(* IEC 61131-3 sources: plc-patterns-examples/listings/BottleFiller, 39 files *)

(* ---- E_ActuatorTarget.st ---- *)
{attribute 'qualified_only'}
{attribute 'strict'}
{attribute 'to_string'}
TYPE E_ActuatorTarget :
(
    None      := 0,     // no move commanded yet; what the outputs do is up to the actuator
    Extended  := 10,
    Retracted := 20
);
END_TYPE

(* ---- E_DeviceSource.st ---- *)
{attribute 'qualified_only'}
{attribute 'strict'}
{attribute 'to_string'}
TYPE E_DeviceSource :
(
    Undefined       := 0,
    FinalHardware   := 1,
    SimilarHardware := 2,
    Simulation      := 3,
    Test            := 4
);
END_TYPE

(* ---- E_FillStep.st ---- *)
{attribute 'qualified_only'}
{attribute 'strict'}
{attribute 'to_string'}
TYPE E_FillStep :
(
    Undefined := 0,
    Idle      := 10,
    Opening   := 20,
    Filling   := 30,
    Closing   := 40,
    Done      := 50,
    Error     := 900
);
END_TYPE

(* ---- E_LineState.st ---- *)
{attribute 'qualified_only'}
{attribute 'strict'}
{attribute 'to_string'}
TYPE E_LineState :
(
    Stopped      := 0,
    Filling      := 10,
    Transferring := 20,
    Faulted      := 900
);
END_TYPE

(* ---- E_OperationState.st ---- *)
{attribute 'qualified_only'}
{attribute 'strict'}
{attribute 'to_string'}
TYPE E_OperationState :
(
    Idle  := 0,     // never started
    Busy  := 1,
    Done  := 2,
    Error := 3
);
END_TYPE

(* ---- E_PickStep.st ---- *)
{attribute 'qualified_only'}
{attribute 'strict'}
{attribute 'to_string'}
TYPE E_PickStep :
(
    Undefined      := 0,
    Idle           := 10,
    LowerToPick    := 20,
    Grip           := 30,
    RaiseWithPart  := 40,
    SlideOut       := 50,
    LowerToPlace   := 60,
    ClampPart      := 65,
    OpenGripper    := 70,
    RaiseEmpty     := 80,
    ReleaseFixture := 85,
    SlideIn        := 90,
    Done           := 100,
    Error          := 900
);
END_TYPE

(* ---- GVL_Hmi.st ---- *)
{attribute 'qualified_only'}
VAR_GLOBAL
    // From the HMI
    StartButton      : BOOL;
    StopButton       : BOOL;
    ResetButton      : BOOL;

    // To the HMI
    LineState        : E_LineState;
    IsStopping       : BOOL;
    FaultText        : STRING;
    NotFinalDevices  : STRING(255);         // every device that isn't the machine's own; empty on the machine
END_VAR

(* ---- GVL_Io.st ---- *)
{attribute 'qualified_only'}
VAR_GLOBAL
    // Filling station
    TankValveCoil  AT %Q* : BOOL;
    TankValveOpen  AT %I* : BOOL;
    DrainValveCoil AT %Q* : BOOL;
    DrainValveOpen AT %I* : BOOL;
    TankLevel      AT %I* : DINT;           // level sensor process data, 0.1 mm
    TankSensorOk   AT %I* : BOOL;           // the sensor's valid bit; see the project document

    // Pick-and-place station
    LiftValve      AT %Q* : BOOL;
    LiftDown       AT %I* : BOOL;
    LiftUp         AT %I* : BOOL;
    SlideOutCoil   AT %Q* : BOOL;
    SlideInCoil    AT %Q* : BOOL;
    SlideOut       AT %I* : BOOL;
    SlideIn        AT %I* : BOOL;
    GripperValve   AT %Q* : BOOL;
    GripperClosed  AT %I* : BOOL;
    GripperOpen    AT %I* : BOOL;
END_VAR

(* ---- GVL_Sim.st ---- *)
{attribute 'qualified_only'}
VAR_GLOBAL
    // Failure hooks for the simulated devices, set from the HMI or a watch
    // window. Each one acts only while its device is simulated.
    TankValveStuck  : BOOL;
    DrainValveStuck : BOOL;
    LiftStuck       : BOOL;
    SlideStuck      : BOOL;
    GripperStuck    : BOOL;
END_VAR

(* ---- GVL_Site.st ---- *)
{attribute 'qualified_only'}
VAR_GLOBAL CONSTANT
    // Edited for each controller; a release never overwrites this list.
    // FinalHardware on the machine. As delivered, everything is simulated.
    TankValveSource  : E_DeviceSource := E_DeviceSource.Simulation;
    DrainValveSource : E_DeviceSource := E_DeviceSource.Simulation;
    TankLevelSource  : E_DeviceSource := E_DeviceSource.Simulation;
    LiftSource       : E_DeviceSource := E_DeviceSource.Simulation;
    SlideSource      : E_DeviceSource := E_DeviceSource.Simulation;
    GripperSource    : E_DeviceSource := E_DeviceSource.Simulation;
    IsOnMachine      : BOOL := FALSE;   // TRUE on the real machine: anything not final is a fault
END_VAR

(* ---- ActuatorBase.st ---- *)
FUNCTION_BLOCK ABSTRACT ActuatorBase IMPLEMENTS I_Actuator, I_Cyclic
VAR
    _Name         : STRING(32);
    _MoveTimeout  : TIME := T#2S;
    _Target       : E_ActuatorTarget;
    _IsInPosition : BOOL;
    _HasFault     : BOOL;
    _FaultText    : STRING(80);
    _MoveTimer    : TON;
    _SettleTimer  : TON;
END_VAR
(*
    ActuatorBase

    The move-and-supervise skeleton shared by every actuator. CyclicLogic() is
    the template: it drives toward the target, checks arrival, supervises the
    move time, goes safe on a fault and lets the actuator settle.

    Derived blocks implement IsWired, DriveOutputs, IsAtPosition and DriveSafe,
    may override SettleTime, and call Configure() from their FB_init.
*)

METHOD PUBLIC FINAL CyclicLogic
// Not wired: report it, touch nothing
IF NOT IsWired() THEN
    _HasFault := TRUE;
    _FaultText := 'I/O not wired';
    RETURN;
END_IF

// Faulted: only the safe outputs, until Reset()
IF _HasFault THEN
    DriveSafe();
    RETURN;
END_IF

// Drive toward the target, and check whether it has arrived
DriveOutputs(Target := _Target);
_IsInPosition := IsAtPosition(Position := _Target);

// Supervise the move: the same rule for every actuator
_MoveTimer(IN := (_Target <> E_ActuatorTarget.None) AND NOT _IsInPosition, PT := _MoveTimeout);
IF _MoveTimer.Q THEN
    _HasFault := TRUE;
    _FaultText := 'Move did not finish in time';
    DriveSafe();
    RETURN;
END_IF

// Let it settle before reporting the position
_SettleTimer(IN := _IsInPosition, PT := SettleTime);

METHOD PROTECTED ABSTRACT IsWired : BOOL

METHOD PROTECTED ABSTRACT DriveOutputs
VAR_INPUT
    Target : E_ActuatorTarget;
END_VAR

METHOD PROTECTED ABSTRACT IsAtPosition : BOOL
VAR_INPUT
    Position : E_ActuatorTarget;
END_VAR

METHOD PROTECTED ABSTRACT DriveSafe

PROPERTY PROTECTED SettleTime : TIME
GET: SettleTime := T#0S;           // most actuators report as soon as the sensor confirms

METHOD PROTECTED Configure
VAR_INPUT
    Name        : STRING(32);
    MoveTimeout : TIME;
END_VAR
_Name := Name;
_MoveTimeout := MoveTimeout;

METHOD PUBLIC Extend
MoveTo(Target := E_ActuatorTarget.Extended);

METHOD PUBLIC Retract
MoveTo(Target := E_ActuatorTarget.Retracted);

METHOD PRIVATE MoveTo
VAR_INPUT
    Target : E_ActuatorTarget;
END_VAR
IF _HasFault OR Target = _Target THEN
    RETURN;                        // faulted: Reset() first. Same target: keep the move running.
END_IF
_Target := Target;
_MoveTimer(IN := FALSE);           // every new move gets the full timeout
_SettleTimer(IN := FALSE);

METHOD PUBLIC Reset
_HasFault := FALSE;
_FaultText := '';
_Target := E_ActuatorTarget.None;
_MoveTimer(IN := FALSE);
_SettleTimer(IN := FALSE);

PROPERTY PUBLIC IsExtended : BOOL
GET: IsExtended := NOT _HasFault AND _Target = E_ActuatorTarget.Extended AND _SettleTimer.Q;

PROPERTY PUBLIC IsRetracted : BOOL
GET: IsRetracted := NOT _HasFault AND _Target = E_ActuatorTarget.Retracted AND _SettleTimer.Q;

PROPERTY PUBLIC HasFault : BOOL
GET: HasFault := _HasFault;

PROPERTY PUBLIC FaultText : STRING
GET: FaultText := _FaultText;

PROPERTY PUBLIC Name : STRING
GET: Name := _Name;

(* ---- ActuatorRouter.st ---- *)
FUNCTION_BLOCK ActuatorRouter IMPLEMENTS I_Actuator, I_Cyclic
VAR
    _Name   : STRING(32);
    _Source : E_DeviceSource;
    _Chosen : I_Actuator;
END_VAR
(*
    ActuatorRouter

    One I_Actuator in front of up to four candidates, chosen once by the
    site setting. Only the chosen candidate is run. A source with no
    candidate (0) is never at either end, and reports a fault.
*)

METHOD FB_init : BOOL
VAR_INPUT
    bInitRetains    : BOOL;
    bInCopyCode     : BOOL;
    Name            : STRING(32);
    Source          : E_DeviceSource;
    FinalHardware   : I_Actuator;
    SimilarHardware : I_Actuator;
    Simulation      : I_Actuator;
    Test            : I_Actuator;
END_VAR
_Name := Name;
_Source := Source;
CASE Source OF
    E_DeviceSource.FinalHardware:   _Chosen := FinalHardware;
    E_DeviceSource.SimilarHardware: _Chosen := SimilarHardware;
    E_DeviceSource.Simulation:      _Chosen := Simulation;
    E_DeviceSource.Test:            _Chosen := Test;
END_CASE

METHOD PUBLIC CyclicLogic
VAR
    Cyclic : I_Cyclic;
END_VAR
IF _Chosen <> 0 AND_THEN __QUERYINTERFACE(_Chosen, Cyclic) THEN
    Cyclic.CyclicLogic();              // only the chosen candidate runs
END_IF

METHOD PUBLIC Extend
IF _Chosen <> 0 THEN
    _Chosen.Extend();
END_IF

METHOD PUBLIC Retract
IF _Chosen <> 0 THEN
    _Chosen.Retract();
END_IF

METHOD PUBLIC Reset
IF _Chosen <> 0 THEN
    _Chosen.Reset();
END_IF

PROPERTY PUBLIC IsExtended : BOOL
GET: IsExtended := _Chosen <> 0 AND_THEN _Chosen.IsExtended;

PROPERTY PUBLIC IsRetracted : BOOL
GET: IsRetracted := _Chosen <> 0 AND_THEN _Chosen.IsRetracted;

PROPERTY PUBLIC Name : STRING
GET: Name := _Name;

PROPERTY PUBLIC HasFault : BOOL
GET: HasFault := _Chosen = 0 OR_ELSE _Chosen.HasFault;

PROPERTY PUBLIC FaultText : STRING
GET:
IF _Chosen = 0 THEN
    FaultText := 'No device for this source';
ELSE
    FaultText := _Chosen.FaultText;
END_IF

PROPERTY PUBLIC Source : E_DeviceSource
GET: Source := _Source;

(* ---- DoubleSolenoidCylinder.st ---- *)
FUNCTION_BLOCK DoubleSolenoidCylinder EXTENDS ActuatorBase
VAR
    _ExtendCoil      : REFERENCE TO BOOL;
    _RetractCoil     : REFERENCE TO BOOL;
    _ExtendedSensor  : REFERENCE TO BOOL;
    _RetractedSensor : REFERENCE TO BOOL;
END_VAR
(*
    DoubleSolenoidCylinder

    One coil per direction. With both coils off, the valve holds the cylinder
    where it is. An end sensor at each end.
*)

METHOD FB_init : BOOL
VAR_INPUT
    bInitRetains    : BOOL;
    bInCopyCode     : BOOL;
    Name            : STRING(32);
    MoveTimeout     : TIME;
    ExtendCoil      : REFERENCE TO BOOL;
    RetractCoil     : REFERENCE TO BOOL;
    ExtendedSensor  : REFERENCE TO BOOL;
    RetractedSensor : REFERENCE TO BOOL;
END_VAR
_ExtendCoil REF= ExtendCoil;
_RetractCoil REF= RetractCoil;
_ExtendedSensor REF= ExtendedSensor;
_RetractedSensor REF= RetractedSensor;
Configure(Name := Name, MoveTimeout := MoveTimeout);

METHOD PROTECTED IsWired : BOOL
IsWired := __ISVALIDREF(_ExtendCoil) AND __ISVALIDREF(_RetractCoil)
       AND __ISVALIDREF(_ExtendedSensor) AND __ISVALIDREF(_RetractedSensor);

METHOD PROTECTED DriveOutputs
VAR_INPUT
    Target : E_ActuatorTarget;
END_VAR
_ExtendCoil := Target = E_ActuatorTarget.Extended;
_RetractCoil := Target = E_ActuatorTarget.Retracted;  // None: both off, so it holds

METHOD PROTECTED IsAtPosition : BOOL
VAR_INPUT
    Position : E_ActuatorTarget;
END_VAR
CASE Position OF
    E_ActuatorTarget.Extended:
        IsAtPosition := _ExtendedSensor AND NOT _RetractedSensor;
    E_ActuatorTarget.Retracted:
        IsAtPosition := _RetractedSensor AND NOT _ExtendedSensor;
ELSE
    IsAtPosition := FALSE;
END_CASE

METHOD PROTECTED DriveSafe
_ExtendCoil := FALSE;                               // both off: the cylinder stays where it is
_RetractCoil := FALSE;

(* ---- DrainTankCommand.st ---- *)
FUNCTION_BLOCK DrainTankCommand IMPLEMENTS I_Command
VAR CONSTANT
    EmptyLevel : REAL := 2.0;          // percent
END_VAR
VAR
    _DrainValve   : I_FillValve;
    _Level        : I_LevelSensor;
    _Clock        : I_Clock;
    _Timeout      : LTIME;
    _StartedAt    : LTIME;
    _State        : E_OperationState;
    _FaultText    : STRING;
    _IsConfigured : BOOL;
END_VAR
(*
    DrainTankCommand

    Opens the drain valve until the tank reads empty. Ends in Error if the
    level sensor is invalid, the valve faults, or the tank isn't empty
    within the timeout. Every ending closes the drain valve.
*)

METHOD FB_init : BOOL
VAR_INPUT
    bInitRetains : BOOL;
    bInCopyCode  : BOOL;
    DrainValve   : I_FillValve;     // any on/off valve with feedback fits this contract
    Level        : I_LevelSensor;
    Clock        : I_Clock;
    Timeout      : LTIME;
END_VAR
_DrainValve := DrainValve;
_Level := Level;
_Clock := Clock;
_Timeout := Timeout;
_IsConfigured := DrainValve <> 0 AND Level <> 0 AND Clock <> 0;

METHOD PUBLIC Start
IF _State = E_OperationState.Busy THEN
    RETURN;
END_IF
IF NOT _IsConfigured THEN
    _State := E_OperationState.Error;
    _FaultText := 'Drain command not wired';
    RETURN;
END_IF
_StartedAt := _Clock.Now;
_FaultText := '';
_State := E_OperationState.Busy;
_DrainValve.Open();

METHOD PUBLIC CyclicLogic
IF _State <> E_OperationState.Busy THEN
    RETURN;
END_IF

IF NOT _Level.IsValid THEN
    Finish(Outcome := E_OperationState.Error, Text := 'Level sensor invalid');
ELSIF _DrainValve.HasFault THEN
    Finish(Outcome := E_OperationState.Error, Text := _DrainValve.FaultText);
ELSIF _Level.Level <= EmptyLevel THEN
    Finish(Outcome := E_OperationState.Done, Text := '');
ELSIF _Clock.Now - _StartedAt >= _Timeout THEN
    Finish(Outcome := E_OperationState.Error, Text := 'Tank did not empty in time');
END_IF

METHOD PUBLIC Abort
IF _State = E_OperationState.Busy THEN
    Finish(Outcome := E_OperationState.Error, Text := 'Aborted');
END_IF

METHOD PRIVATE Finish
VAR_INPUT
    Outcome : E_OperationState;
    Text    : STRING;
END_VAR
_DrainValve.Close();                 // every ending, good or bad, leaves the drain closed
_State := Outcome;
_FaultText := Text;

PROPERTY PUBLIC Name : STRING
GET: Name := 'Drain tank';

PROPERTY PUBLIC State : E_OperationState
GET: State := _State;

PROPERTY PUBLIC FaultText : STRING
GET: FaultText := _FaultText;

(* ---- EquipmentGroup.st ---- *)
FUNCTION_BLOCK EquipmentGroup IMPLEMENTS I_Diagnosable, I_Resettable
VAR CONSTANT
    MaxChildren : DINT := 16;
END_VAR
VAR
    _Name        : STRING(32);
    _Children    : ARRAY[0..MaxChildren - 1] OF I_Diagnosable;
    _Resettables : ARRAY[0..MaxChildren - 1] OF I_Resettable;
    _Count       : DINT;
END_VAR
(*
    EquipmentGroup

    A named group of devices or other groups, behind the same interfaces
    as one device. It has a fault while any child has one, and reports
    the first faulted child's text, prefixed with that child's name.
    Reset() resets every child that implements I_Resettable.
    AddChild() is called while wiring, before the group is first asked.
*)

METHOD FB_init : BOOL
VAR_INPUT
    bInitRetains : BOOL;
    bInCopyCode  : BOOL;
    Name         : STRING(32);
END_VAR
_Name := Name;

METHOD PUBLIC AddChild : BOOL
VAR_INPUT
    Child : I_Diagnosable;
END_VAR
VAR
    Me         : I_Diagnosable;
    Resettable : I_Resettable;
    i          : DINT;
END_VAR
Me := THIS^;
IF Child = 0 OR Child = Me OR _Count >= MaxChildren THEN
    AddChild := FALSE;
    RETURN;
END_IF
FOR i := 0 TO _Count - 1 DO           // the same child only once
    IF _Children[i] = Child THEN
        AddChild := FALSE;
        RETURN;
    END_IF
END_FOR
_Children[_Count] := Child;
IF __QUERYINTERFACE(Child, Resettable) THEN
    _Resettables[_Count] := Resettable;
END_IF
_Count := _Count + 1;
AddChild := TRUE;

METHOD PUBLIC Reset
VAR
    i : DINT;
END_VAR
FOR i := 0 TO _Count - 1 DO
    IF _Resettables[i] <> 0 THEN
        _Resettables[i].Reset();
    END_IF
END_FOR

METHOD PRIVATE FirstFaultIndex : DINT
VAR
    i : DINT;
END_VAR
FOR i := 0 TO _Count - 1 DO
    IF _Children[i].HasFault THEN
        FirstFaultIndex := i;
        RETURN;
    END_IF
END_FOR
FirstFaultIndex := _Count;            // no child has a fault

METHOD PRIVATE DescribeFault : STRING
VAR_INPUT
    Index : DINT;
END_VAR
IF Index < _Count THEN
    DescribeFault := CONCAT(CONCAT(_Children[Index].Name, ': '), _Children[Index].FaultText);
END_IF

PROPERTY PUBLIC Name : STRING
GET: Name := _Name;

PROPERTY PUBLIC HasFault : BOOL
GET: HasFault := FirstFaultIndex() < _Count;

PROPERTY PUBLIC FaultText : STRING
GET: FaultText := DescribeFault(Index := FirstFaultIndex());

PROPERTY PUBLIC ChildCount : DINT
GET: ChildCount := _Count;

(* ---- FakeClock.st ---- *)
FUNCTION_BLOCK FakeClock IMPLEMENTS I_Clock
VAR
    _Now : LTIME;
END_VAR
(*
    FakeClock

    Stands still until the test moves it.
*)

METHOD PUBLIC Advance
VAR_INPUT
    Duration : LTIME;
END_VAR
_Now := _Now + Duration;

PROPERTY PUBLIC Now : LTIME
GET: Now := _Now;

(* ---- FakeEquipmentModule.st ---- *)
FUNCTION_BLOCK FakeEquipmentModule IMPLEMENTS I_EquipmentModule, I_Resettable
VAR
    _Name        : STRING(32);
    _IsCycleDone : BOOL;
    _HasFault    : BOOL;
    _StartCount  : DINT;
    _ResetCount  : DINT;
END_VAR
(*
    FakeEquipmentModule

    Test double for I_EquipmentModule. Counts the cycles it was asked for
    and the resets it received. A requested cycle finishes when the test
    calls FinishCycle(); a fault is reported while the test sets one.
*)

METHOD FB_init : BOOL
VAR_INPUT
    bInitRetains : BOOL;
    bInCopyCode  : BOOL;
    Name         : STRING(32);
END_VAR
_Name := Name;

METHOD PUBLIC StartCycle
_StartCount := _StartCount + 1;
_IsCycleDone := FALSE;

METHOD PUBLIC Reset
_ResetCount := _ResetCount + 1;

METHOD PUBLIC FinishCycle
_IsCycleDone := TRUE;

METHOD PUBLIC SetFault
VAR_INPUT
    IsActive : BOOL;
END_VAR
_HasFault := IsActive;

PROPERTY PUBLIC Name : STRING
GET: Name := _Name;

PROPERTY PUBLIC HasFault : BOOL
GET: HasFault := _HasFault;

PROPERTY PUBLIC FaultText : STRING
GET:
IF _HasFault THEN
    FaultText := 'Simulated fault';
ELSE
    FaultText := '';
END_IF

PROPERTY PUBLIC IsCycleDone : BOOL
GET: IsCycleDone := _IsCycleDone;

PROPERTY PUBLIC StartCount : DINT
GET: StartCount := _StartCount;

PROPERTY PUBLIC ResetCount : DINT
GET: ResetCount := _ResetCount;

(* ---- FieldbusLevelSensor.st ---- *)
FUNCTION_BLOCK FieldbusLevelSensor IMPLEMENTS I_LevelSensor
VAR
    _FieldbusLevel     : REFERENCE TO DINT;
    _IsCommunicationOk : REFERENCE TO BOOL;
    _TankHeight        : REAL;
    _IsConfigured      : BOOL;
END_VAR
(* FieldbusLevelSensor: a level sensor that reports its reading over a fieldbus, in 0.1 mm. *)

METHOD FB_init : BOOL
VAR_INPUT
    bInitRetains      : BOOL;
    bInCopyCode       : BOOL;
    FieldbusLevel     : REFERENCE TO DINT;   // process data from the sensor, 0.1 mm
    IsCommunicationOk : REFERENCE TO BOOL;
    TankHeight        : REAL;                // mm
END_VAR
_FieldbusLevel REF= FieldbusLevel;
_IsCommunicationOk REF= IsCommunicationOk;
_TankHeight := TankHeight;
_IsConfigured := __ISVALIDREF(FieldbusLevel) AND __ISVALIDREF(IsCommunicationOk) AND TankHeight > 0.0;

PROPERTY PUBLIC IsValid : BOOL
GET: IsValid := _IsConfigured AND_THEN _IsCommunicationOk;

PROPERTY PUBLIC Level : REAL
GET:
IF IsValid THEN
    Level := LIMIT(0.0, DINT_TO_REAL(_FieldbusLevel) / 10.0 / _TankHeight * 100.0, 100.0);
ELSE
    Level := 0.0;
END_IF

(* ---- FillingModule.st ---- *)
FUNCTION_BLOCK FillingModule EXTENDS ModuleGroup IMPLEMENTS I_EquipmentModule
VAR
    _Fill             : REFERENCE TO FillSequence;
    _Dose             : I_Command;
    _IsCycleRequested : BOOL;
    _IsFilling        : BOOL;
    _IsDosing         : BOOL;
    _HasDoseFault     : BOOL;
    _DoseFault        : STRING;
    _IsConfigured     : BOOL;
END_VAR
(*
    FillingModule

    The filling station. One cycle measures one dose: the fill sequence
    fills the dosing tank to its target level, then the dose command
    drains it into the bottle below. Runs both before its valves. It has
    a fault while a valve has one, the fill sequence has stopped with an
    error, or the last dose ended in Error; Reset() clears all three.
*)

METHOD FB_init : BOOL
VAR_INPUT
    bInitRetains : BOOL;
    bInCopyCode  : BOOL;
    Name         : STRING(32);                  // for EquipmentGroup
    Fill         : REFERENCE TO FillSequence;
    Dose         : I_Command;
END_VAR
_Fill REF= Fill;
_Dose := Dose;
_IsConfigured := __ISVALIDREF(Fill) AND Dose <> 0;

METHOD PUBLIC StartCycle
_IsCycleRequested := TRUE;

METHOD PROTECTED BeforeChildren
IF NOT _IsConfigured THEN
    RETURN;
END_IF

// A new cycle starts with the fill, once the station is free
IF _IsCycleRequested AND NOT _IsFilling AND NOT _IsDosing
   AND (_Fill.CurrentStep = E_FillStep.Idle OR _Fill.CurrentStep = E_FillStep.Done) THEN
    _Fill.Start();
    _IsFilling := TRUE;
    _IsCycleRequested := FALSE;
END_IF
_Fill.CyclicLogic();

// The tank is at its level: dose it into the bottle
IF _IsFilling AND _Fill.IsDone THEN
    _IsFilling := FALSE;
    _Dose.Start();
    _IsDosing := TRUE;
END_IF
IF _IsDosing THEN
    _Dose.CyclicLogic();
    IF _Dose.State = E_OperationState.Error THEN
        _HasDoseFault := TRUE;
        _DoseFault := _Dose.FaultText;
        _IsDosing := FALSE;
    ELSIF _Dose.State = E_OperationState.Done THEN
        _IsDosing := FALSE;
    END_IF
END_IF

METHOD PUBLIC Reset
SUPER^.Reset();                                 // the valves
IF NOT _IsConfigured THEN
    RETURN;
END_IF
_Fill.Reset();
IF _IsDosing THEN
    _Dose.Abort();                              // closes the drain valve
END_IF
_IsCycleRequested := FALSE;
_IsFilling := FALSE;
_IsDosing := FALSE;
_HasDoseFault := FALSE;
_DoseFault := '';

PROPERTY PUBLIC IsCycleDone : BOOL
GET:
IsCycleDone := _IsConfigured AND_THEN (NOT _IsCycleRequested AND NOT _IsFilling AND NOT _IsDosing
                                             AND _Dose.State = E_OperationState.Done);

PROPERTY PUBLIC HasFault : BOOL
GET:
IF NOT _IsConfigured THEN
    HasFault := TRUE;
ELSE
    HasFault := SUPER^.HasFault OR _Fill.HasError OR _HasDoseFault;
END_IF

PROPERTY PUBLIC FaultText : STRING
GET:
IF NOT _IsConfigured THEN
    FaultText := 'Filling station not wired';
ELSIF SUPER^.HasFault THEN
    FaultText := SUPER^.FaultText;              // the valve, by name
ELSIF _Fill.HasError THEN
    FaultText := 'Fill stopped; reset to continue';
ELSIF _HasDoseFault THEN
    FaultText := CONCAT('Dose: ', _DoseFault);
ELSE
    FaultText := '';
END_IF

(* ---- FillSequence.st ---- *)
FUNCTION_BLOCK FillSequence
VAR
    _LevelSensor      : I_LevelSensor;
    _FillValve        : I_FillValve;
    _TargetLevel      : REAL := 80.0;
    _CurrentStep      : E_FillStep := E_FillStep.Idle;
    _IsStartRequested : BOOL;
    _IsResetRequested : BOOL;
    _IsConfigured     : BOOL;
END_VAR
(*
    FillSequence

    Opens the fill valve, waits for the target level, closes the valve.
    Talks only to I_LevelSensor and I_FillValve, injected through FB_init.

    Call CyclicLogic() once per cycle. Start() and Reset() are requests,
    seen during the next CyclicLogic() call.
*)

METHOD PUBLIC Start
_IsStartRequested := TRUE;

METHOD PUBLIC Reset
_IsResetRequested := TRUE;

METHOD PUBLIC CyclicLogic
IF NOT _IsConfigured THEN
    _CurrentStep := E_FillStep.Error;   // not wired: fail safe, never call through 0
    RETURN;
END_IF

CASE _CurrentStep OF
    E_FillStep.Idle, E_FillStep.Done:
        IF _IsStartRequested THEN
            _CurrentStep := E_FillStep.Opening;
        END_IF

    E_FillStep.Opening:
        _FillValve.Open();
        IF _FillValve.IsOpen THEN
            _CurrentStep := E_FillStep.Filling;
        ELSIF _FillValve.HasFault THEN
            _CurrentStep := E_FillStep.Error;
        END_IF

    E_FillStep.Filling:
        IF NOT _LevelSensor.IsValid OR _FillValve.HasFault THEN
            _CurrentStep := E_FillStep.Error;
        ELSIF _LevelSensor.Level >= _TargetLevel THEN
            _CurrentStep := E_FillStep.Closing;
        END_IF

    E_FillStep.Closing:
        _FillValve.Close();
        IF _FillValve.IsClosed THEN
            _CurrentStep := E_FillStep.Done;
        ELSIF _FillValve.HasFault THEN
            _CurrentStep := E_FillStep.Error;
        END_IF

    E_FillStep.Error:
        _FillValve.Close();             // the one promise every valve keeps
        IF _IsResetRequested AND _FillValve.IsClosed THEN
            _CurrentStep := E_FillStep.Idle;
        END_IF
END_CASE

_IsStartRequested := FALSE;
_IsResetRequested := FALSE;

PROPERTY PUBLIC TargetLevel : REAL
GET: TargetLevel := _TargetLevel;
SET: _TargetLevel := LIMIT(0.0, TargetLevel, 100.0);

PROPERTY PUBLIC CurrentStep : E_FillStep
GET: CurrentStep := _CurrentStep;

PROPERTY PUBLIC IsBusy : BOOL
GET:
IsBusy := _CurrentStep = E_FillStep.Opening
            OR _CurrentStep = E_FillStep.Filling
            OR _CurrentStep = E_FillStep.Closing;

PROPERTY PUBLIC IsDone : BOOL
GET: IsDone := _CurrentStep = E_FillStep.Done;

PROPERTY PUBLIC HasError : BOOL
GET: HasError := _CurrentStep = E_FillStep.Error;

METHOD FB_init : BOOL
VAR_INPUT
    bInitRetains : BOOL;
    bInCopyCode  : BOOL;
    LevelSensor  : I_LevelSensor;
    FillValve    : I_FillValve;
END_VAR
_LevelSensor := LevelSensor;
_FillValve := FillValve;
_IsConfigured := LevelSensor <> 0 AND FillValve <> 0;   // stored: FB_init's return value is ignored

(* ---- FillValveRouter.st ---- *)
FUNCTION_BLOCK FillValveRouter IMPLEMENTS I_FillValve, I_Cyclic
VAR
    _Name   : STRING(32);
    _Source : E_DeviceSource;
    _Chosen : I_FillValve;
END_VAR
(*
    FillValveRouter

    One I_FillValve in front of up to four candidates. The site setting,
    given once in FB_init, chooses which candidate answers and which one
    is run. A source with no candidate (0) reports a fault and is never
    open.
*)

METHOD FB_init : BOOL
VAR_INPUT
    bInitRetains    : BOOL;
    bInCopyCode     : BOOL;
    Name            : STRING(32);
    Source          : E_DeviceSource;
    FinalHardware   : I_FillValve;
    SimilarHardware : I_FillValve;
    Simulation      : I_FillValve;
    Test            : I_FillValve;
END_VAR
_Name := Name;
_Source := Source;
CASE Source OF
    E_DeviceSource.FinalHardware:   _Chosen := FinalHardware;
    E_DeviceSource.SimilarHardware: _Chosen := SimilarHardware;
    E_DeviceSource.Simulation:      _Chosen := Simulation;
    E_DeviceSource.Test:            _Chosen := Test;
END_CASE

METHOD PUBLIC CyclicLogic
VAR
    Cyclic : I_Cyclic;
END_VAR
IF _Chosen <> 0 AND_THEN __QUERYINTERFACE(_Chosen, Cyclic) THEN
    Cyclic.CyclicLogic();              // only the chosen candidate runs
END_IF

METHOD PUBLIC Open
IF _Chosen <> 0 THEN
    _Chosen.Open();
END_IF

METHOD PUBLIC Close
IF _Chosen <> 0 THEN
    _Chosen.Close();
END_IF

PROPERTY PUBLIC IsOpen : BOOL
GET: IsOpen := _Chosen <> 0 AND_THEN _Chosen.IsOpen;

PROPERTY PUBLIC IsClosed : BOOL
GET: IsClosed := _Chosen <> 0 AND_THEN _Chosen.IsClosed;

PROPERTY PUBLIC Name : STRING
GET: Name := _Name;

PROPERTY PUBLIC HasFault : BOOL
GET: HasFault := _Chosen = 0 OR_ELSE _Chosen.HasFault;

PROPERTY PUBLIC FaultText : STRING
GET:
IF _Chosen = 0 THEN
    FaultText := 'No device for this source';
ELSE
    FaultText := _Chosen.FaultText;
END_IF

PROPERTY PUBLIC Source : E_DeviceSource
GET: Source := _Source;

(* ---- LevelSensorRouter.st ---- *)
FUNCTION_BLOCK LevelSensorRouter IMPLEMENTS I_LevelSensor, I_Cyclic
VAR
    _Name   : STRING(32);
    _Source : E_DeviceSource;
    _Chosen : I_LevelSensor;
END_VAR
(*
    LevelSensorRouter

    One I_LevelSensor in front of up to four candidates, chosen once by
    the site setting. A source with no candidate (0) is never valid.
*)

METHOD FB_init : BOOL
VAR_INPUT
    bInitRetains    : BOOL;
    bInCopyCode     : BOOL;
    Name            : STRING(32);
    Source          : E_DeviceSource;
    FinalHardware   : I_LevelSensor;
    SimilarHardware : I_LevelSensor;
    Simulation      : I_LevelSensor;
    Test            : I_LevelSensor;
END_VAR
_Name := Name;
_Source := Source;
CASE Source OF
    E_DeviceSource.FinalHardware:   _Chosen := FinalHardware;
    E_DeviceSource.SimilarHardware: _Chosen := SimilarHardware;
    E_DeviceSource.Simulation:      _Chosen := Simulation;
    E_DeviceSource.Test:            _Chosen := Test;
END_CASE

METHOD PUBLIC CyclicLogic
VAR
    Cyclic : I_Cyclic;
END_VAR
IF _Chosen <> 0 AND_THEN __QUERYINTERFACE(_Chosen, Cyclic) THEN
    Cyclic.CyclicLogic();              // only the chosen candidate runs
END_IF

PROPERTY PUBLIC Level : REAL
GET:
IF _Chosen <> 0 THEN
    Level := _Chosen.Level;
ELSE
    Level := 0.0;
END_IF

PROPERTY PUBLIC IsValid : BOOL
GET: IsValid := _Chosen <> 0 AND_THEN _Chosen.IsValid;

PROPERTY PUBLIC Name : STRING
GET: Name := _Name;

PROPERTY PUBLIC Source : E_DeviceSource
GET: Source := _Source;

(* ---- LineModule.st ---- *)
FUNCTION_BLOCK LineModule EXTENDS ModuleGroup
VAR
    _Filler           : I_EquipmentModule;
    _Transfer         : I_EquipmentModule;
    _State            : E_LineState;
    _IsStartRequested : BOOL;
    _IsStopping       : BOOL;
    _IsConfigured     : BOOL;
END_VAR
(*
    LineModule

    The machine module. Fills a bottle, moves it out, and repeats until
    stopped. Commands its two stations in BeforeChildren(), before they
    run in the same scan.

    Start() starts the line. Stop() lets the bottle in progress finish.
    A fault anywhere in the tree stops commanding and shows Faulted; once
    the tree no longer reports a fault, the line is Stopped and waits for
    Start(). Reset(), inherited, resets the whole tree.
*)

METHOD FB_init : BOOL
VAR_INPUT
    bInitRetains : BOOL;
    bInCopyCode  : BOOL;
    Name         : STRING(32);                  // for EquipmentGroup
    Filler       : I_EquipmentModule;
    Transfer     : I_EquipmentModule;
END_VAR
_Filler := Filler;
_Transfer := Transfer;
_IsConfigured := Filler <> 0 AND Transfer <> 0;

METHOD PUBLIC Start
_IsStartRequested := TRUE;
_IsStopping := FALSE;                           // a start cancels a stop that hasn't been taken yet

METHOD PUBLIC Stop
IF _State <> E_LineState.Stopped THEN
    _IsStopping := TRUE;                        // taken when the bottle is out
END_IF

METHOD PROTECTED BeforeChildren
IF NOT _IsConfigured THEN
    _State := E_LineState.Faulted;
    RETURN;
END_IF

// A fault anywhere in the tree: command nothing
IF HasFault THEN
    _State := E_LineState.Faulted;
    _IsStopping := FALSE;
    _IsStartRequested := FALSE;
    RETURN;
END_IF

CASE _State OF
    E_LineState.Stopped:
        IF _IsStartRequested THEN
            _Filler.StartCycle();
            _State := E_LineState.Filling;
        END_IF

    E_LineState.Filling:
        IF _Filler.IsCycleDone THEN
            _Transfer.StartCycle();
            _State := E_LineState.Transferring;
        END_IF

    E_LineState.Transferring:
        IF _Transfer.IsCycleDone THEN
            IF _IsStopping THEN
                _IsStopping := FALSE;
                _State := E_LineState.Stopped;
            ELSE
                _Filler.StartCycle();           // the next bottle
                _State := E_LineState.Filling;
            END_IF
        END_IF

    E_LineState.Faulted:
        _State := E_LineState.Stopped;          // no fault any more; wait for Start
END_CASE

_IsStartRequested := FALSE;

PROPERTY PUBLIC State : E_LineState
GET: State := _State;

PROPERTY PUBLIC IsStopping : BOOL
GET: IsStopping := _IsStopping;

(* ---- LineRunsStopsAndFaultsTest.st ---- *)
FUNCTION_BLOCK LineRunsStopsAndFaultsTest EXTENDS TestBase
VAR
    _Filler   : FakeEquipmentModule(Name := 'Filling');
    _Transfer : FakeEquipmentModule(Name := 'Pick and place');
    _Line     : LineModule(Name := 'Line 1', Filler := _Filler, Transfer := _Transfer);
    _IsWired  : BOOL;
END_VAR
(*
    LineRunsStopsAndFaultsTest

    The line fills, then transfers, and repeats; a stop is taken at the end
    of the bottle; a fault stops all commands until it clears, and the line
    then waits for a new start.
*)

METHOD PUBLIC Run
// The fakes are children too, so the line sees their faults and resets them
_IsWired := _Line.AddChild(Child := _Filler) AND _Line.AddChild(Child := _Transfer);
Check(_IsWired, 'both stations added');

// Power-up: stopped, nothing commanded
_Line.CyclicLogic();
Check(_Line.State = E_LineState.Stopped AND _Filler.StartCount = 0, 'stopped at power-up');

// Start: one bottle is filled
_Line.Start();
_Line.CyclicLogic();
Check(_Line.State = E_LineState.Filling AND _Filler.StartCount = 1, 'start fills a bottle');

// The fill is not done yet: the line waits
_Line.CyclicLogic();
Check(_Line.State = E_LineState.Filling AND _Transfer.StartCount = 0, 'waits for the fill');

// The fill is done: the bottle is moved out
_Filler.FinishCycle();
_Line.CyclicLogic();
Check(_Line.State = E_LineState.Transferring AND _Transfer.StartCount = 1, 'then transfers');

// The transfer is done: the next bottle is filled
_Transfer.FinishCycle();
_Line.CyclicLogic();
Check(_Line.State = E_LineState.Filling AND _Filler.StartCount = 2, 'then fills the next bottle');

// Stop during a fill: the bottle is finished first
_Line.Stop();
_Line.CyclicLogic();
Check(_Line.State = E_LineState.Filling AND _Line.IsStopping, 'stop waits for the bottle');
_Filler.FinishCycle();
_Line.CyclicLogic();
Check(_Line.State = E_LineState.Transferring, 'the bottle is still moved out');
_Transfer.FinishCycle();
_Line.CyclicLogic();
Check(_Line.State = E_LineState.Stopped AND _Filler.StartCount = 2, 'then stops, with no new fill');

// A fault: nothing is commanded, not even a start
_Line.Start();
_Filler.SetFault(IsActive := TRUE);
_Line.CyclicLogic();
Check(_Line.State = E_LineState.Faulted AND _Filler.StartCount = 2, 'a fault blocks the start');

// Reset reaches every station
_Line.Reset();
Check(_Filler.ResetCount = 1 AND _Transfer.ResetCount = 1, 'reset reaches both stations');

// The fault clears: stopped, and waiting for a new start
_Filler.SetFault(IsActive := FALSE);
_Line.CyclicLogic();
Check(_Line.State = E_LineState.Stopped AND _Filler.StartCount = 2, 'stopped after the fault, no restart');

(* ---- ModuleGroup.st ---- *)
FUNCTION_BLOCK ModuleGroup EXTENDS EquipmentGroup IMPLEMENTS I_Cyclic
VAR
    _Cyclics : ARRAY[0..MaxChildren - 1] OF I_Cyclic;
END_VAR
(*
    ModuleGroup

    An EquipmentGroup that also runs its children: one CyclicLogic() call
    runs every child that implements I_Cyclic, in the order they were
    added, between this module's own BeforeChildren() and AfterChildren().
    A station with logic of its own extends it and overrides the hooks.
*)

METHOD PUBLIC AddChild : BOOL
VAR_INPUT
    Child : I_Diagnosable;
END_VAR
VAR
    Cyclic : I_Cyclic;
END_VAR
IF NOT SUPER^.AddChild(Child := Child) THEN
    AddChild := FALSE;
    RETURN;
END_IF
IF __QUERYINTERFACE(Child, Cyclic) THEN
    _Cyclics[_Count - 1] := Cyclic;   // the slot SUPER^.AddChild() just filled
END_IF
AddChild := TRUE;

METHOD PUBLIC FINAL CyclicLogic
VAR
    i : DINT;
END_VAR
BeforeChildren();
FOR i := 0 TO _Count - 1 DO
    IF _Cyclics[i] <> 0 THEN
        _Cyclics[i].CyclicLogic();
    END_IF
END_FOR
AfterChildren();

METHOD PROTECTED BeforeChildren      // decide what the children should do this scan

METHOD PROTECTED AfterChildren       // read what they reported this scan

(* ---- PickAndPlaceModule.st ---- *)
FUNCTION_BLOCK PickAndPlaceModule EXTENDS ModuleGroup IMPLEMENTS I_EquipmentModule
VAR
    _Sequence         : REFERENCE TO PickAndPlaceSequence;
    _IsCycleRequested : BOOL;
    _IsConfigured     : BOOL;
END_VAR
(*
    PickAndPlaceModule

    The pick-and-place station. Runs its PickAndPlaceSequence, then its
    actuators. One StartCycle() moves one bottle from the filler to the
    outfeed. It has a fault while the sequence reports one, which includes
    every actuator's; Reset() resets both.
*)

METHOD FB_init : BOOL
VAR_INPUT
    bInitRetains : BOOL;
    bInCopyCode  : BOOL;
    Name         : STRING(32);                  // for EquipmentGroup
    Sequence     : REFERENCE TO PickAndPlaceSequence;
END_VAR
_Sequence REF= Sequence;
_IsConfigured := __ISVALIDREF(Sequence);

METHOD PUBLIC StartCycle
_IsCycleRequested := TRUE;

METHOD PROTECTED BeforeChildren
IF NOT _IsConfigured THEN
    RETURN;
END_IF
IF _IsCycleRequested
   AND (_Sequence.CurrentStep = E_PickStep.Idle OR _Sequence.CurrentStep = E_PickStep.Done) THEN
    _Sequence.Start();
    _IsCycleRequested := FALSE;
END_IF
_Sequence.CyclicLogic();                        // the sequence decides; the actuators move after it

METHOD PUBLIC Reset
SUPER^.Reset();                                 // the actuators
IF _IsConfigured THEN
    _Sequence.Reset();
END_IF
_IsCycleRequested := FALSE;

PROPERTY PUBLIC IsCycleDone : BOOL
GET: IsCycleDone := _IsConfigured AND_THEN (NOT _IsCycleRequested AND _Sequence.CurrentStep = E_PickStep.Done);

PROPERTY PUBLIC HasFault : BOOL
GET:
IF NOT _IsConfigured THEN
    HasFault := TRUE;
ELSE
    HasFault := SUPER^.HasFault OR _Sequence.HasFault;
END_IF

PROPERTY PUBLIC FaultText : STRING
GET:
IF NOT _IsConfigured THEN
    FaultText := 'Pick and place not wired';
ELSIF SUPER^.HasFault THEN
    FaultText := SUPER^.FaultText;              // the actuator, by name
ELSIF _Sequence.HasFault THEN
    FaultText := _Sequence.FaultText;
ELSE
    FaultText := '';
END_IF

(* ---- PickAndPlaceSequence.st ---- *)
FUNCTION_BLOCK PickAndPlaceSequence
VAR
    _Lift            : I_Actuator;
    _Slide           : I_Actuator;
    _Gripper         : I_Actuator;
    _CurrentStep      : E_PickStep;
    _FaultText        : STRING;
    _IsStartRequested : BOOL;
    _IsResetRequested : BOOL;
    _IsConfigured     : BOOL;
END_VAR
(*
    PickAndPlaceSequence

    Picks a part, slides across, places it and slides back. Moves three
    I_Actuator, injected through FB_init, and never knows what kind each
    one is.

    Call CyclicLogic() once per cycle. Start() and Reset() are requests,
    seen during the next CyclicLogic() call. After a reset it returns home the way a cycle ends:
    lift up, then slide in.
*)

METHOD FB_init : BOOL
VAR_INPUT
    bInitRetains : BOOL;
    bInCopyCode  : BOOL;
    Lift         : I_Actuator;      // extended = down
    Slide        : I_Actuator;      // extended = over the place position
    Gripper      : I_Actuator;      // extended = closed
END_VAR
_Lift := Lift;
_Slide := Slide;
_Gripper := Gripper;
_IsConfigured := Lift <> 0 AND Slide <> 0 AND Gripper <> 0;

METHOD PUBLIC Start
_IsStartRequested := TRUE;

METHOD PUBLIC Reset
_IsResetRequested := TRUE;

METHOD PUBLIC CyclicLogic
IF NOT _IsConfigured THEN
    _CurrentStep := E_PickStep.Error;      // not wired: never call through 0
    _FaultText := 'Pick and place not wired';
    RETURN;
END_IF

CASE _CurrentStep OF
    E_PickStep.Undefined:
        _CurrentStep := E_PickStep.Idle;

    E_PickStep.Idle, E_PickStep.Done:
        IF _IsStartRequested THEN
            _CurrentStep := E_PickStep.LowerToPick;
        END_IF

    E_PickStep.LowerToPick:   ExtendThen(Actuator := _Lift, NextStep := E_PickStep.Grip);
    E_PickStep.Grip:          ExtendThen(Actuator := _Gripper, NextStep := E_PickStep.RaiseWithPart);
    E_PickStep.RaiseWithPart: RetractThen(Actuator := _Lift, NextStep := E_PickStep.SlideOut);
    E_PickStep.SlideOut:      ExtendThen(Actuator := _Slide, NextStep := E_PickStep.LowerToPlace);
    E_PickStep.LowerToPlace:  ExtendThen(Actuator := _Lift, NextStep := E_PickStep.OpenGripper);
    E_PickStep.OpenGripper:   RetractThen(Actuator := _Gripper, NextStep := E_PickStep.RaiseEmpty);
    E_PickStep.RaiseEmpty:    RetractThen(Actuator := _Lift, NextStep := E_PickStep.SlideIn);
    E_PickStep.SlideIn:       RetractThen(Actuator := _Slide, NextStep := E_PickStep.Done);

    E_PickStep.Error:
        IF _IsResetRequested THEN
            _Lift.Reset(); _Slide.Reset(); _Gripper.Reset();
            _FaultText := '';
            _CurrentStep := E_PickStep.RaiseEmpty;   // go home the way a cycle ends
        END_IF
END_CASE

_IsStartRequested := FALSE;
_IsResetRequested := FALSE;

METHOD PRIVATE ExtendThen
VAR_INPUT
    Actuator : I_Actuator;
    NextStep : E_PickStep;
END_VAR
Actuator.Extend();
IF Actuator.IsExtended THEN
    _CurrentStep := NextStep;
ELSIF Actuator.HasFault THEN
    Fail(Actuator := Actuator);
END_IF

METHOD PRIVATE RetractThen
VAR_INPUT
    Actuator : I_Actuator;
    NextStep : E_PickStep;
END_VAR
Actuator.Retract();
IF Actuator.IsRetracted THEN
    _CurrentStep := NextStep;
ELSIF Actuator.HasFault THEN
    Fail(Actuator := Actuator);
END_IF

METHOD PRIVATE Fail
VAR_INPUT
    Actuator : I_Actuator;
END_VAR
_FaultText := CONCAT(CONCAT(Actuator.Name, ': '), Actuator.FaultText);
_CurrentStep := E_PickStep.Error;

PROPERTY PUBLIC CurrentStep : E_PickStep
GET: CurrentStep := _CurrentStep;

PROPERTY PUBLIC IsBusy : BOOL
GET:
IsBusy := _CurrentStep <> E_PickStep.Undefined AND _CurrentStep <> E_PickStep.Idle
            AND _CurrentStep <> E_PickStep.Done AND _CurrentStep <> E_PickStep.Error;

PROPERTY PUBLIC HasFault : BOOL
GET:
IF _IsConfigured THEN
    HasFault := _Lift.HasFault OR _Slide.HasFault OR _Gripper.HasFault;
END_IF
HasFault := HasFault OR _CurrentStep = E_PickStep.Error;

PROPERTY PUBLIC FaultText : STRING
GET: FaultText := _FaultText;

(* ---- SimulatedActuator.st ---- *)
FUNCTION_BLOCK SimulatedActuator EXTENDS ActuatorBase
VAR
    _TravelTime   : TIME;
    _DrivenTarget : E_ActuatorTarget;
    _Travel       : TON;
    _IsStuck      : BOOL;
END_VAR
(*
    SimulatedActuator

    Stands in for a cylinder or gripper with end sensors. Reaches the
    commanded end TravelTime after the move starts. The supervision is
    ActuatorBase's, unchanged, so a move that never arrives faults exactly
    as a real one would. SetStuck() stops it moving. Has no I/O.
*)

METHOD FB_init : BOOL
VAR_INPUT
    bInitRetains : BOOL;
    bInCopyCode  : BOOL;
    Name         : STRING(32);
    MoveTimeout  : TIME;
    TravelTime   : TIME;
END_VAR
_TravelTime := TravelTime;
Configure(Name := Name, MoveTimeout := MoveTimeout);

METHOD PUBLIC SetStuck
VAR_INPUT
    IsStuck : BOOL;
END_VAR
_IsStuck := IsStuck;

METHOD PROTECTED IsWired : BOOL
IsWired := TRUE;                                    // nothing to wire

METHOD PROTECTED DriveOutputs
VAR_INPUT
    Target : E_ActuatorTarget;
END_VAR
IF Target <> _DrivenTarget THEN
    _DrivenTarget := Target;
    _Travel(IN := FALSE);                           // a new move starts from the beginning
END_IF
_Travel(IN := Target <> E_ActuatorTarget.None AND NOT _IsStuck, PT := _TravelTime);

METHOD PROTECTED IsAtPosition : BOOL
VAR_INPUT
    Position : E_ActuatorTarget;
END_VAR
IsAtPosition := Position <> E_ActuatorTarget.None AND Position = _DrivenTarget AND _Travel.Q;

METHOD PROTECTED DriveSafe
_Travel(IN := FALSE);

(* ---- SimulatedValve.st ---- *)
FUNCTION_BLOCK SimulatedValve IMPLEMENTS I_FillValve, I_Cyclic
VAR
    _Name         : STRING(32);
    _Clock        : I_Clock;
    _TravelTime   : LTIME;
    _IsCommanded  : BOOL;              // TRUE: open requested
    _IsStuck      : BOOL;
    _IsAtOpen     : BOOL;
    _IsAtClosed   : BOOL := TRUE;
    _MoveStart    : LTIME;
    _IsMoving     : BOOL;
    _IsConfigured : BOOL;
END_VAR
(*
    SimulatedValve

    Stands in for a valve with position feedback. Reaches the commanded
    position after TravelTime, with neither end reported while it moves.
    SetStuck() makes it stop answering commands, as a sticking valve does.
    Has no I/O.
*)

METHOD FB_init : BOOL
VAR_INPUT
    bInitRetains : BOOL;
    bInCopyCode  : BOOL;
    Name         : STRING(32);
    Clock        : I_Clock;
    TravelTime   : LTIME;
END_VAR
_Name := Name;
_Clock := Clock;
_TravelTime := TravelTime;
_IsConfigured := Clock <> 0;

METHOD PUBLIC Open
_IsCommanded := TRUE;

METHOD PUBLIC Close
_IsCommanded := FALSE;

METHOD PUBLIC SetStuck
VAR_INPUT
    IsStuck : BOOL;
END_VAR
_IsStuck := IsStuck;

METHOD PUBLIC CyclicLogic
IF NOT _IsConfigured OR _IsStuck THEN
    RETURN;
END_IF
IF _IsCommanded <> _IsAtOpen AND NOT _IsMoving THEN
    _IsMoving := TRUE;                 // a new command: leave the end position
    _MoveStart := _Clock.Now;
    _IsAtOpen := FALSE;
    _IsAtClosed := FALSE;
END_IF
IF _IsMoving AND_THEN _Clock.Now - _MoveStart >= _TravelTime THEN
    _IsMoving := FALSE;
    _IsAtOpen := _IsCommanded;
    _IsAtClosed := NOT _IsCommanded;
END_IF

PROPERTY PUBLIC IsOpen : BOOL
GET: IsOpen := _IsAtOpen;

PROPERTY PUBLIC IsClosed : BOOL
GET: IsClosed := _IsAtClosed;

PROPERTY PUBLIC Name : STRING
GET: Name := _Name;

PROPERTY PUBLIC HasFault : BOOL
GET: HasFault := NOT _IsConfigured;

PROPERTY PUBLIC FaultText : STRING
GET: FaultText := SEL(_IsConfigured, 'Simulated valve has no clock', '');

(* ---- SimulatedValveTakesItsTravelTimeTest.st ---- *)
FUNCTION_BLOCK SimulatedValveTakesItsTravelTimeTest EXTENDS TestBase
VAR
    _Clock : FakeClock;
    _Valve : SimulatedValve(Name := 'Test valve', Clock := _Clock, TravelTime := LTIME#400MS);
END_VAR
(*
    SimulatedValveTakesItsTravelTimeTest

    The simulated valve reports neither end while it travels, reaches open
    after its travel time, and doesn't move at all while stuck.
*)

METHOD PUBLIC Run
Check(_Valve.IsClosed AND NOT _Valve.IsOpen, 'it starts closed');

_Valve.Open();
_Valve.CyclicLogic();
Check(NOT _Valve.IsClosed AND NOT _Valve.IsOpen, 'it reports neither end while it travels');

_Clock.Advance(Duration := LTIME#399MS);
_Valve.CyclicLogic();
Check(NOT _Valve.IsOpen, 'it is not open before its travel time');

_Clock.Advance(Duration := LTIME#1MS);
_Valve.CyclicLogic();
Check(_Valve.IsOpen, 'it is open after its travel time');

_Valve.SetStuck(IsStuck := TRUE);
_Valve.Close();
_Clock.Advance(Duration := LTIME#1S);
_Valve.CyclicLogic();
Check(_Valve.IsOpen, 'a stuck valve ignores Close()');

(* ---- SimulationCheck.st ---- *)
FUNCTION_BLOCK SimulationCheck IMPLEMENTS I_Diagnosable
VAR
    _IsOnMachine    : BOOL;
    _NotFinalCount  : DINT;
    _NotFinalNames  : STRING(255);
END_VAR
(*
    SimulationCheck

    Told, while wiring, the name and source of every routed device. Lists
    every device that isn't FinalHardware, for the HMI and the event log.
    On a controller whose site is the machine itself, each of them is a
    fault.
*)

METHOD FB_init : BOOL
VAR_INPUT
    bInitRetains : BOOL;
    bInCopyCode  : BOOL;
    IsOnMachine  : BOOL;
END_VAR
_IsOnMachine := IsOnMachine;

METHOD PUBLIC AddDevice : BOOL
VAR_INPUT
    Name   : STRING(32);
    Source : E_DeviceSource;
END_VAR
AddDevice := TRUE;
IF Source = E_DeviceSource.FinalHardware THEN
    RETURN;
END_IF
_NotFinalCount := _NotFinalCount + 1;
IF _NotFinalCount = 1 THEN
    _NotFinalNames := Name;
ELSE
    _NotFinalNames := CONCAT(CONCAT(_NotFinalNames, ', '), Name);
END_IF

PROPERTY PUBLIC Name : STRING
GET: Name := 'Device sources';

PROPERTY PUBLIC HasFault : BOOL
GET: HasFault := _IsOnMachine AND _NotFinalCount > 0;

PROPERTY PUBLIC FaultText : STRING
GET:
IF HasFault THEN
    FaultText := CONCAT('Not final hardware: ', _NotFinalNames);
ELSE
    FaultText := '';
END_IF

PROPERTY PUBLIC NotFinalDevices : STRING(255)
GET: NotFinalDevices := _NotFinalNames;

PROPERTY PUBLIC NotFinalCount : DINT
GET: NotFinalCount := _NotFinalCount;

(* ---- SimulationCheckTest.st ---- *)
FUNCTION_BLOCK SimulationCheckTest EXTENDS TestBase
VAR
    _OnDesk    : SimulationCheck(IsOnMachine := FALSE);
    _OnMachine : SimulationCheck(IsOnMachine := TRUE);
    _Ok        : BOOL;
END_VAR
(*
    SimulationCheckTest

    Every device that isn't final hardware is listed; only on the machine
    is that a fault.
*)

METHOD PUBLIC Run
_Ok := _OnDesk.AddDevice(Name := 'Tank valve', Source := E_DeviceSource.Simulation);
_Ok := _OnDesk.AddDevice(Name := 'Lift', Source := E_DeviceSource.FinalHardware) AND _Ok;
_Ok := _OnDesk.AddDevice(Name := 'Tank level', Source := E_DeviceSource.SimilarHardware) AND _Ok;
Check(_Ok, 'every device is accepted');
Check(_OnDesk.NotFinalCount = 2 AND _OnDesk.NotFinalDevices = 'Tank valve, Tank level',
      'the devices that are not final hardware are listed');
Check(NOT _OnDesk.HasFault, 'on a desk, that is not a fault');

_OnMachine.AddDevice(Name := 'Lift', Source := E_DeviceSource.FinalHardware);
Check(NOT _OnMachine.HasFault, 'on the machine, final hardware is no fault');
_OnMachine.AddDevice(Name := 'Tank valve', Source := E_DeviceSource.Simulation);
Check(_OnMachine.HasFault, 'on the machine, a simulated device is a fault');

(* ---- SingleSolenoidCylinder.st ---- *)
FUNCTION_BLOCK SingleSolenoidCylinder EXTENDS ActuatorBase
VAR
    _Solenoid        : REFERENCE TO BOOL;
    _ExtendedSensor  : REFERENCE TO BOOL;
    _RetractedSensor : REFERENCE TO BOOL;
END_VAR
(*
    SingleSolenoidCylinder

    One solenoid with spring return: energized extends, de-energized retracts.
    An end sensor at each end.
*)

METHOD FB_init : BOOL
VAR_INPUT
    bInitRetains    : BOOL;
    bInCopyCode     : BOOL;
    Name            : STRING(32);
    MoveTimeout     : TIME;
    Solenoid        : REFERENCE TO BOOL;
    ExtendedSensor  : REFERENCE TO BOOL;
    RetractedSensor : REFERENCE TO BOOL;
END_VAR
_Solenoid REF= Solenoid;
_ExtendedSensor REF= ExtendedSensor;
_RetractedSensor REF= RetractedSensor;
Configure(Name := Name, MoveTimeout := MoveTimeout);

METHOD PROTECTED IsWired : BOOL
IsWired := __ISVALIDREF(_Solenoid) AND __ISVALIDREF(_ExtendedSensor) AND __ISVALIDREF(_RetractedSensor);

METHOD PROTECTED DriveOutputs
VAR_INPUT
    Target : E_ActuatorTarget;
END_VAR
_Solenoid := Target = E_ActuatorTarget.Extended;   // anything else: the spring retracts it

METHOD PROTECTED IsAtPosition : BOOL
VAR_INPUT
    Position : E_ActuatorTarget;
END_VAR
CASE Position OF
    E_ActuatorTarget.Extended:
        IsAtPosition := _ExtendedSensor AND NOT _RetractedSensor;
    E_ActuatorTarget.Retracted:
        IsAtPosition := _RetractedSensor AND NOT _ExtendedSensor;
ELSE
    IsAtPosition := FALSE;
END_CASE

METHOD PROTECTED DriveSafe
_Solenoid := FALSE;                                 // the spring takes it to the retracted end

(* ---- SolenoidValve.st ---- *)
FUNCTION_BLOCK SolenoidValve IMPLEMENTS I_FillValve, I_Resettable, I_Cyclic
VAR
    _Name          : STRING(32) := 'Solenoid valve';
    _Output        : REFERENCE TO BOOL;
    _OpenFeedback  : REFERENCE TO BOOL;
    _FaultDelay    : TIME;
    _Command       : BOOL;
    _MismatchTimer : TON;
    _IsConfigured  : BOOL;
END_VAR
(*
    SolenoidValve

    Drives one solenoid valve and checks its open-feedback switch. A fault
    is reported while the feedback has disagreed with the command for
    longer than FaultDelay. Name can be set while wiring.
*)

METHOD FB_init : BOOL
VAR_INPUT
    bInitRetains : BOOL;
    bInCopyCode  : BOOL;
    Output       : REFERENCE TO BOOL;
    OpenFeedback : REFERENCE TO BOOL;
    FaultDelay   : TIME;
END_VAR
_Output REF= Output;
_OpenFeedback REF= OpenFeedback;
_FaultDelay := FaultDelay;
_IsConfigured := __ISVALIDREF(Output) AND __ISVALIDREF(OpenFeedback);

METHOD PUBLIC Open
_Command := TRUE;

METHOD PUBLIC Close
_Command := FALSE;

METHOD PUBLIC CyclicLogic
IF NOT _IsConfigured THEN
    RETURN;
END_IF
_Output := _Command;
_MismatchTimer(IN := _Command XOR _OpenFeedback, PT := _FaultDelay);

METHOD PUBLIC Reset
_MismatchTimer(IN := FALSE);                        // supervise again from now

PROPERTY PUBLIC IsOpen : BOOL
GET: IsOpen := _IsConfigured AND_THEN (_Command AND _OpenFeedback);

PROPERTY PUBLIC IsClosed : BOOL
GET: IsClosed := _IsConfigured AND_THEN NOT (_Command OR _OpenFeedback);

PROPERTY PUBLIC HasFault : BOOL
GET: HasFault := NOT _IsConfigured OR _MismatchTimer.Q;

PROPERTY PUBLIC FaultText : STRING
GET:
IF NOT _IsConfigured THEN
    FaultText := 'I/O not wired';
ELSIF _MismatchTimer.Q THEN
    FaultText := 'No feedback';
ELSE
    FaultText := '';
END_IF

PROPERTY PUBLIC Name : STRING
GET: Name := _Name;
SET: _Name := Name;

(* ---- TankModel.st ---- *)
FUNCTION_BLOCK TankModel IMPLEMENTS I_LevelSensor, I_Cyclic
VAR
    _Inflow       : I_FillValve;
    _Outflow      : I_FillValve;
    _Clock        : I_Clock;
    _FillRate     : REAL;              // percent per second, inflow valve open
    _DrainRate    : REAL;              // percent per second, outflow valve open
    _Level        : REAL;
    _LastNow      : LTIME;
    _IsStarted    : BOOL;
    _IsConfigured : BOOL;
END_VAR
(*
    TankModel

    A simulated tank: the level rises while the inflow valve is open and
    falls while the outflow valve is open. Reads both through
    I_FillValve, so it works with simulated and real valves alike.
*)

METHOD FB_init : BOOL
VAR_INPUT
    bInitRetains : BOOL;
    bInCopyCode  : BOOL;
    Inflow       : I_FillValve;
    Outflow      : I_FillValve;
    Clock        : I_Clock;
    FillRate     : REAL;
    DrainRate    : REAL;
    StartLevel   : REAL;
END_VAR
_Inflow := Inflow;
_Outflow := Outflow;
_Clock := Clock;
_FillRate := FillRate;
_DrainRate := DrainRate;
_Level := StartLevel;
_IsConfigured := Inflow <> 0 AND Outflow <> 0 AND Clock <> 0;

METHOD PUBLIC CyclicLogic
VAR
    Now     : LTIME;
    Seconds : REAL;
END_VAR
IF NOT _IsConfigured THEN
    RETURN;
END_IF
Now := _Clock.Now;
IF NOT _IsStarted THEN
    _IsStarted := TRUE;
    _LastNow := Now;
    RETURN;
END_IF
Seconds := LREAL_TO_REAL(LTIME_TO_LREAL(Now - _LastNow) / 1.0E9);   // LTIME counts nanoseconds
_LastNow := Now;
IF _Inflow.IsOpen THEN
    _Level := _Level + _FillRate * Seconds;
END_IF
IF _Outflow.IsOpen THEN
    _Level := _Level - _DrainRate * Seconds;
END_IF
_Level := LIMIT(0.0, _Level, 100.0);

PROPERTY PUBLIC Level : REAL
GET: Level := _Level;

PROPERTY PUBLIC IsValid : BOOL
GET: IsValid := _IsConfigured;

(* ---- TaskClock.st ---- *)
FUNCTION_BLOCK TaskClock IMPLEMENTS I_Clock
VAR
    _CycleTime : LTIME;
    _Now       : LTIME;
END_VAR
(*
    TaskClock

    Advances by the task's cycle time on every CyclicLogic() call. Call it
    once per scan, first, before anything that reads Now.
*)

METHOD FB_init : BOOL
VAR_INPUT
    bInitRetains : BOOL;
    bInCopyCode  : BOOL;
    CycleTime    : LTIME;
END_VAR
_CycleTime := CycleTime;

METHOD PUBLIC CyclicLogic
_Now := _Now + _CycleTime;

PROPERTY PUBLIC Now : LTIME
GET: Now := _Now;

(* ---- TestBase.st ---- *)
FUNCTION_BLOCK ABSTRACT TestBase
VAR
    _CheckCount  : INT;
    _FailedCount : INT;
    _LastFailure : STRING(255);
END_VAR
(*
    TestBase

    Shared bookkeeping for framework-free tests. A derived test implements
    Run() and calls Check() for everything it wants to verify.
*)

METHOD PUBLIC ABSTRACT Run

METHOD PROTECTED Check
VAR_INPUT
    Condition : BOOL;
    Message   : STRING(255);    // what should be true, not what went wrong
END_VAR
_CheckCount := _CheckCount + 1;
IF NOT Condition THEN
    _FailedCount := _FailedCount + 1;
    _LastFailure := Message;
END_IF

PROPERTY PUBLIC HasPassed : BOOL
GET: HasPassed := _CheckCount > 0 AND _FailedCount = 0;

PROPERTY PUBLIC FailedCount : INT
GET: FailedCount := _FailedCount;

PROPERTY PUBLIC LastFailure : STRING(255)
GET: LastFailure := _LastFailure;

(* ---- MAIN.st ---- *)
PROGRAM MAIN
VAR
    Clock         : TaskClock(CycleTime := LTIME#10MS);

    // Filling station: every candidate is declared; the routers choose
    RealTankValve  : SolenoidValve(Output := GVL_Io.TankValveCoil,
                                   OpenFeedback := GVL_Io.TankValveOpen,
                                   FaultDelay := T#2S);
    SimTankValve   : SimulatedValve(Name := 'Tank valve', Clock := Clock, TravelTime := LTIME#400MS);
    TankValve      : FillValveRouter(Name := 'Tank valve', Source := GVL_Site.TankValveSource,
                                     FinalHardware := RealTankValve, SimilarHardware := 0,
                                     Simulation := SimTankValve, Test := 0);

    RealDrainValve : SolenoidValve(Output := GVL_Io.DrainValveCoil,
                                   OpenFeedback := GVL_Io.DrainValveOpen,
                                   FaultDelay := T#2S);
    SimDrainValve  : SimulatedValve(Name := 'Drain valve', Clock := Clock, TravelTime := LTIME#400MS);
    DrainValve     : FillValveRouter(Name := 'Drain valve', Source := GVL_Site.DrainValveSource,
                                     FinalHardware := RealDrainValve, SimilarHardware := 0,
                                     Simulation := SimDrainValve, Test := 0);

    SimTank        : TankModel(Inflow := TankValve, Outflow := DrainValve, Clock := Clock,
                               FillRate := 20.0, DrainRate := 25.0, StartLevel := 0.0);
    RealLevel      : FieldbusLevelSensor(FieldbusLevel := GVL_Io.TankLevel,
                                         IsCommunicationOk := GVL_Io.TankSensorOk,
                                         TankHeight := 300.0);          // the dosing tank, mm
    TankLevel      : LevelSensorRouter(Name := 'Tank level', Source := GVL_Site.TankLevelSource,
                                       FinalHardware := RealLevel, SimilarHardware := 0,
                                       Simulation := SimTank, Test := 0);

    // Pick-and-place station
    RealLift       : SingleSolenoidCylinder(Name := 'Lift', MoveTimeout := T#1S,
                                            Solenoid := GVL_Io.LiftValve,
                                            ExtendedSensor := GVL_Io.LiftDown,
                                            RetractedSensor := GVL_Io.LiftUp);
    SimLift        : SimulatedActuator(Name := 'Lift', MoveTimeout := T#1S, TravelTime := T#400MS);
    LiftCylinder   : ActuatorRouter(Name := 'Lift', Source := GVL_Site.LiftSource,
                                    FinalHardware := RealLift, SimilarHardware := 0,
                                    Simulation := SimLift, Test := 0);

    RealSlide      : DoubleSolenoidCylinder(Name := 'Slide', MoveTimeout := T#2S,
                                            ExtendCoil := GVL_Io.SlideOutCoil,
                                            RetractCoil := GVL_Io.SlideInCoil,
                                            ExtendedSensor := GVL_Io.SlideOut,
                                            RetractedSensor := GVL_Io.SlideIn);
    SimSlide       : SimulatedActuator(Name := 'Slide', MoveTimeout := T#2S, TravelTime := T#800MS);
    SlideCylinder  : ActuatorRouter(Name := 'Slide', Source := GVL_Site.SlideSource,
                                    FinalHardware := RealSlide, SimilarHardware := 0,
                                    Simulation := SimSlide, Test := 0);

    RealGripper    : Gripper(Name := 'Gripper', MoveTimeout := T#500MS,
                             Solenoid := GVL_Io.GripperValve,
                             ExtendedSensor := GVL_Io.GripperClosed,
                             RetractedSensor := GVL_Io.GripperOpen);
    SimGripper     : SimulatedActuator(Name := 'Gripper', MoveTimeout := T#500MS, TravelTime := T#150MS);
    PartGripper    : ActuatorRouter(Name := 'Gripper', Source := GVL_Site.GripperSource,
                                    FinalHardware := RealGripper, SimilarHardware := 0,
                                    Simulation := SimGripper, Test := 0);

    // The operations, unchanged from their pages
    TankFill       : FillSequence(LevelSensor := TankLevel, FillValve := TankValve);
    Dose           : DrainTankCommand(DrainValve := DrainValve, Level := TankLevel,
                                      Clock := Clock, Timeout := LTIME#30S);
    PickPlace      : PickAndPlaceSequence(Lift := LiftCylinder, Slide := SlideCylinder,
                                          Gripper := PartGripper);

    // The tree
    Sources        : SimulationCheck(IsOnMachine := GVL_Site.IsOnMachine);
    Filling        : FillingModule(Name := 'Filling', Fill := TankFill, Dose := Dose);
    PickAndPlace   : PickAndPlaceModule(Name := 'Pick and place', Sequence := PickPlace);
    Line           : LineModule(Name := 'Line 1', Filler := Filling, Transfer := PickAndPlace);

    StartEdge      : R_TRIG;
    StopEdge       : R_TRIG;
    ResetEdge      : R_TRIG;
    Wired          : BOOL;
    WiredOk        : BOOL;
END_VAR

// Build the tree once, and tell the check where every device comes from
IF NOT Wired THEN
    Wired := TRUE;
    WiredOk := Filling.AddChild(Child := TankValve);
    WiredOk := Filling.AddChild(Child := DrainValve) AND WiredOk;
    WiredOk := PickAndPlace.AddChild(Child := LiftCylinder) AND WiredOk;
    WiredOk := PickAndPlace.AddChild(Child := SlideCylinder) AND WiredOk;
    WiredOk := PickAndPlace.AddChild(Child := PartGripper) AND WiredOk;
    WiredOk := Line.AddChild(Child := Sources) AND WiredOk;
    WiredOk := Line.AddChild(Child := Filling) AND WiredOk;
    WiredOk := Line.AddChild(Child := PickAndPlace) AND WiredOk;

    WiredOk := Sources.AddDevice(Name := TankValve.Name, Source := TankValve.Source) AND WiredOk;
    WiredOk := Sources.AddDevice(Name := DrainValve.Name, Source := DrainValve.Source) AND WiredOk;
    WiredOk := Sources.AddDevice(Name := TankLevel.Name, Source := TankLevel.Source) AND WiredOk;
    WiredOk := Sources.AddDevice(Name := LiftCylinder.Name, Source := LiftCylinder.Source) AND WiredOk;
    WiredOk := Sources.AddDevice(Name := SlideCylinder.Name, Source := SlideCylinder.Source) AND WiredOk;
    WiredOk := Sources.AddDevice(Name := PartGripper.Name, Source := PartGripper.Source) AND WiredOk;
    GVL_Hmi.NotFinalDevices := Sources.NotFinalDevices;
END_IF

// Failure hooks act only on a simulated device
IF TankValve.Source = E_DeviceSource.Simulation THEN
    SimTankValve.SetStuck(IsStuck := GVL_Sim.TankValveStuck);
END_IF
IF DrainValve.Source = E_DeviceSource.Simulation THEN
    SimDrainValve.SetStuck(IsStuck := GVL_Sim.DrainValveStuck);
END_IF
IF LiftCylinder.Source = E_DeviceSource.Simulation THEN
    SimLift.SetStuck(IsStuck := GVL_Sim.LiftStuck);
END_IF
IF SlideCylinder.Source = E_DeviceSource.Simulation THEN
    SimSlide.SetStuck(IsStuck := GVL_Sim.SlideStuck);
END_IF
IF PartGripper.Source = E_DeviceSource.Simulation THEN
    SimGripper.SetStuck(IsStuck := GVL_Sim.GripperStuck);
END_IF

// Operator commands
StartEdge(CLK := GVL_Hmi.StartButton);
StopEdge(CLK := GVL_Hmi.StopButton);
ResetEdge(CLK := GVL_Hmi.ResetButton);
IF StartEdge.Q AND WiredOk THEN
    Line.Start();
END_IF
IF StopEdge.Q THEN
    Line.Stop();
END_IF
IF ResetEdge.Q THEN
    Line.Reset();
END_IF

Clock.CyclicLogic();                            // first: everything below reads its time
TankLevel.CyclicLogic();                        // runs the tank model only when it's the chosen level
Line.CyclicLogic();                             // the line, then each station, then its devices

GVL_Hmi.LineState := Line.State;
GVL_Hmi.IsStopping := Line.IsStopping;
GVL_Hmi.FaultText := Line.FaultText;

(* ---- TestMain.st ---- *)
PROGRAM TestMain
VAR
    LineTest    : LineRunsStopsAndFaultsTest;
    ValveTest   : SimulatedValveTakesItsTravelTimeTest;
    CheckTest   : SimulationCheckTest;
    HasRun      : BOOL;
    AllPassed   : BOOL;
    FailedCount : INT;
END_VAR

// Each test runs once, on the first scan. None of them touches the machine's
// instances or its I/O. Read AllPassed, FailedCount and each test's
// LastFailure in a watch window.
IF NOT HasRun THEN
    HasRun := TRUE;
    LineTest.Run();
    ValveTest.Run();
    CheckTest.Run();
    AllPassed := LineTest.HasPassed AND ValveTest.HasPassed AND CheckTest.HasPassed;
    FailedCount := LineTest.FailedCount + ValveTest.FailedCount + CheckTest.FailedCount;
END_IF
